// TIA Portal V20 export
// export: Created 2026-10-12T05:42:30.1522252Z, ExportSetting WithDefaults, DisplayName Totally Integrated Automation Portal, DisplayVersion V20, DisplayName TIA Portal Openness, DisplayVersion V20, DisplayName TIA Portal Teamcenter Gateway, DisplayVersion V20, DisplayName TIA Portal Version Control Interface, DisplayVersion V20, DisplayName SINAMICS Startdrive Advanced, DisplayVersion V20 SP1 Update 2, DisplayName SINAMICS Startdrive G110M, G120, G120C, G120D, G120P, G115D, DisplayVersion V20 SP1 Update 2, DisplayName SINAMICS Startdrive G130, G150, S120, S150, SINAMICS MV, G220, S200, S210, DisplayVersion V20 SP1 Update 2, DisplayName STEP 7 Professional, DisplayVersion V20, DisplayName STEP 7 Safety, DisplayVersion V20, DisplayName WinCC Basic/Comfort/Advanced, DisplayVersion V20, DisplayName WinCC Professional, DisplayVersion V20, DisplayName WinCC Unified, DisplayVersion V20
FUNCTION "FRK_AccessPolicyBoot" : Void   // FC59, SCL
{ S7_Optimized_Access := 'TRUE' }
VERSION : 0.1
// stored: AutoNumber true, IsIECCheckEnabled false, SetENOAutomatically false, UDAEnableTagReadback false
   VAR_INPUT
      Startup : Bool;
      Root : Bool;
      Scope : String;
   END_VAR
   VAR_IN_OUT
      Access : "FRK_Access";
   END_VAR
   VAR_TEMP
      Index : Int;
      FreeSlot : Int;
   END_VAR
BEGIN

   IF NOT #Startup THEN
       RETURN;
   END_IF;
   #Access.PolicySlot := 0;
   #Access.PolicyLost := FALSE;
   #Access.PolicyLossAlarm := 0;
   #Access.UserLossAlarm := 0;
   IF NOT #Root THEN
       RETURN;
   END_IF;
   #FreeSlot := 0;
   FOR #Index := 1 TO 1 DO
       IF "FRK_AccessPolicies".Rows[#Index].Scope = #Scope THEN
           IF #Access.PolicySlot <> 0 THEN
               #Access.PolicyLost := TRUE;
           ELSE
               #Access.PolicySlot := #Index;
           END_IF;
       ELSIF #FreeSlot = 0 AND NOT "FRK_AccessPolicies".Rows[#Index].Initialized AND "FRK_AccessPolicies".Rows[#Index].Scope = '' AND "FRK_AccessPolicies".Rows[#Index].SchemaVersion = 0 AND "FRK_AccessPolicies".Rows[#Index].Generation = 0 AND "FRK_AccessPolicies".Rows[#Index].Checksum = DWORD#0 THEN
           #FreeSlot := #Index;
       END_IF;
   END_FOR;
   IF #Access.PolicySlot > 0 THEN
       IF NOT #Access.PolicyLost AND "FRK_AccessPolicyValid"(Image := "FRK_AccessPolicies".Rows[#Access.PolicySlot]) THEN
           #Access.Policy := "FRK_AccessPolicies".Rows[#Access.PolicySlot].Policy;
       ELSE
           #Access.PolicyLost := TRUE;
       END_IF;
   ELSIF #FreeSlot > 0 THEN
       #Access.PolicySlot := #FreeSlot;
       "FRK_AccessPolicySave"(Access := #Access,
                              Scope := #Scope);
   ELSE
       #Access.PolicyLost := TRUE;
   END_IF;
   IF #Access.PolicyLost THEN
       // Do not silently reopen actions after losing commissioned policy.
       #Access.Policy := "FRK_AccessStorage".EmptyPolicy;
       FOR #Index := 0 TO 11 DO
           #Access.Policy.Required[#Index] := 4;
       END_FOR;
   END_IF;
END_FUNCTION
